FUNCTION_BLOCK OutputHanding (* Composite Function Block Type *)
  (* Standard: 61499-2 *)
  (* Version 0.0, 7/2/2026, template *)
  PACKAGE Main;
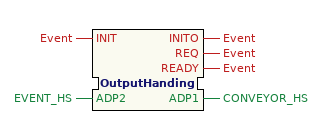
  EVENT_INPUT
    INIT; (* Initialization Request *)
  END_EVENT
  EVENT_OUTPUT
    INITO; (* Initialization Confirm *)
    REQ; (* Execution Confirmation *)
    READY;
  END_EVENT
  SOCKETS
    ADP2 : EVENT_HS;
  END_SOCKETS
  PLUGS
    ADP1 : CONVEYOR_HS;
  END_PLUGS
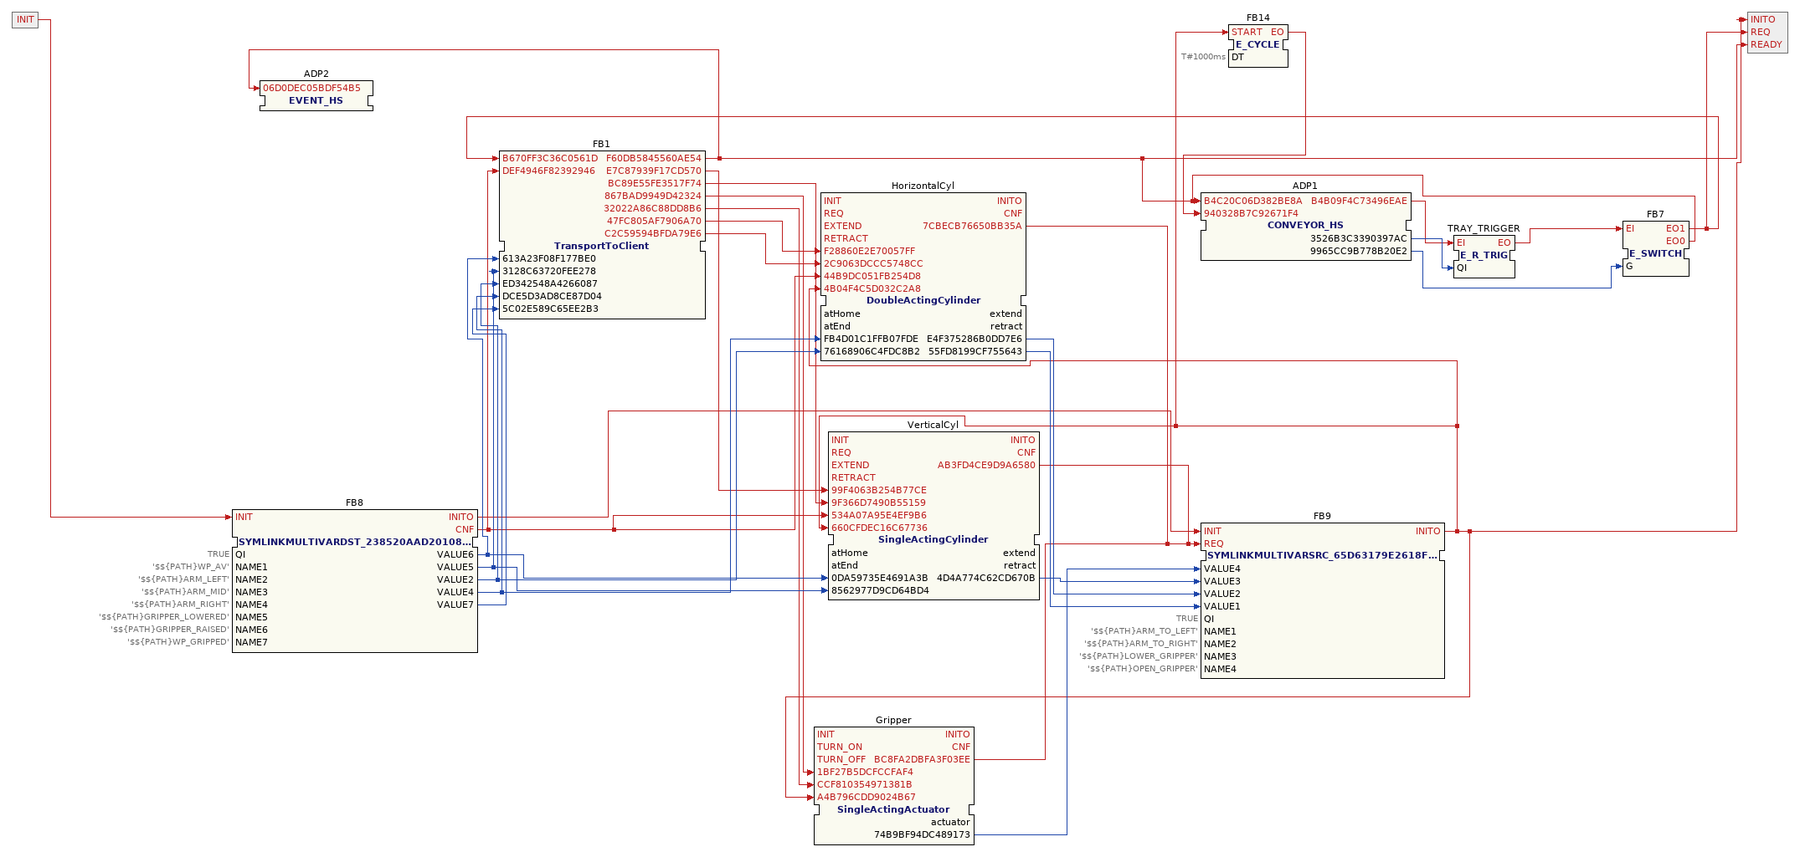
  FBS
    FB1 : TransportToClient;
    HorizontalCyl : DoubleActingCylinder;
    VerticalCyl : SingleActingCylinder;
    Gripper : SingleActingActuator;
    FB14 : E_CYCLE(DT := T#1000ms);
    TRAY_TRIGGER : E_R_TRIG;
    FB7 : E_SWITCH;
    FB8 : SYMLINKMULTIVARDST_238520AAD20108C65(QI := TRUE, NAME1 := '$${PATH}WP_AV', NAME2 := '$${PATH}ARM_LEFT', NAME3 := '$${PATH}ARM_MID', NAME4 := '$${PATH}ARM_RIGHT', NAME5 := '$${PATH}GRIPPER_LOWERED', NAME6 := '$${PATH}GRIPPER_RAISED', NAME7 := '$${PATH}WP_GRIPPED'); {SET_ATTRIBUTE(Configuration.GenericFBType.InterfaceParams, Runtime.System#I:=7;VALUE${I$}:BOOL,BOOL,BOOL,BOOL,BOOL,BOOL,BOOL)}
    FB9 : SYMLINKMULTIVARSRC_65D63179E2618F5E(QI := TRUE, NAME1 := '$${PATH}ARM_TO_LEFT', NAME2 := '$${PATH}ARM_TO_RIGHT', NAME3 := '$${PATH}LOWER_GRIPPER', NAME4 := '$${PATH}OPEN_GRIPPER'); {SET_ATTRIBUTE(Configuration.GenericFBType.InterfaceParams, Runtime.System#I:=5;VALUE${I$}:BOOL,BOOL,BOOL,BOOL,BOOL)}
  END_FBS
  EVENT_CONNECTIONS
    INIT TO FB8.INIT;
    FB1.F60DB5845560AE54 TO ADP2.06D0DEC05BDF54B5;
    FB1.F60DB5845560AE54 TO READY;
    FB1.F60DB5845560AE54 TO ADP1.B4C20C06D382BE8A;
    FB7.EO1 TO FB1.B670FF3C36C0561D;
    FB7.EO1 TO REQ;
    FB8.INITO TO FB9.INIT;
    FB1.E7C87939F17CD570 TO VerticalCyl.99F4063B254B77CE;
    FB1.BC89E55FE3517F74 TO VerticalCyl.9F366D7490B55159;
    FB1.867BAD9949D42324 TO Gripper.1BF27B5DCFCCFAF4;
    FB1.32022A86C88DD8B6 TO Gripper.CCF810354971381B;
    FB1.47FC805AF7906A70 TO HorizontalCyl.F28860E2E70057FF;
    FB1.C2C59594BFDA79E6 TO HorizontalCyl.2C9063DCCC5748CC;
    FB9.INITO TO FB14.START;
    FB14.EO TO ADP1.940328B7C92671F4;
    ADP1.B4B09F4C73496EAE TO TRAY_TRIGGER.EI;
    TRAY_TRIGGER.EO TO FB7.EI;
    FB7.EO0 TO ADP1.B4C20C06D382BE8A;
    FB9.INITO TO INITO;
    FB8.CNF TO FB1.DEF4946F82392946;
    FB8.CNF TO HorizontalCyl.44B9DC051FB254D8;
    FB8.CNF TO VerticalCyl.534A07A95E4EF9B6;
    HorizontalCyl.7CBECB76650BB35A TO FB9.REQ;
    VerticalCyl.AB3FD4CE9D9A6580 TO FB9.REQ;
    Gripper.BC8FA2DBFA3F03EE TO FB9.REQ;
    FB9.INITO TO HorizontalCyl.4B04F4C5D032C2A8;
    FB9.INITO TO VerticalCyl.660CFDEC16C67736;
    FB9.INITO TO Gripper.A4B796CDD9024B67;
  END_CONNECTIONS
  DATA_CONNECTIONS
    FB8.VALUE6 TO FB1.613A23F08F177BE0;
    FB8.VALUE5 TO FB1.3128C63720FEE278;
    FB8.VALUE2 TO FB1.ED342548A4266087;
    FB8.VALUE4 TO FB1.DCE5D3AD8CE87D04;
    FB8.VALUE7 TO FB1.5C02E589C65EE2B3;
    ADP1.3526B3C3390397AC TO TRAY_TRIGGER.QI;
    ADP1.9965CC9B778B20E2 TO FB7.G;
    Gripper.74B9BF94DC489173 TO FB9.VALUE4;
    VerticalCyl.4D4A774C62CD670B TO FB9.VALUE3;
    HorizontalCyl.E4F375286B0DD7E6 TO FB9.VALUE2;
    HorizontalCyl.55FD8199CF755643 TO FB9.VALUE1;
    FB8.VALUE6 TO VerticalCyl.0DA59735E4691A3B;
    FB8.VALUE5 TO VerticalCyl.8562977D9CD64BD4;
    FB8.VALUE4 TO HorizontalCyl.FB4D01C1FFB07FDE;
    FB8.VALUE2 TO HorizontalCyl.76168906C4FDC8B2;
  END_CONNECTIONS
END_FUNCTION_BLOCK
